(* IEC 61131-3 sources: Elmo_Master/Lasal_PRG/Welcon8Axis_EtherCAT_Test_With_RobotAxis/Network/TCPComNet, 1 file *)

(* ---- ONE_TCPComNet_Table.st ---- *)
#define OBJECTS_CONFIG

#include "..\..\Class\DataManager\DataManager.h"
//Define part of class DataManagerFIFO
#define MEMORY_Mark_DataMngFiFo    8
#include <.\lsl_st_mt.h>
#include "..\..\Class\TCPCommunication\TCPCommunication.h"
#include "..\..\Class\TCPCommunication\SalamanderDelay.h"

FUNCTION GLOBAL TAB ONE_TCPComNet
-1$UINT, 0$UINT,
0$UINT, 0$UINT,

15$UDINT,
TO_UDINT(916194998), "_CheckSum", 1$UINT, 0$UINT, 1$UINT,
TO_UDINT(3238142347), "_SigTCPComReceive", 1$UINT, 1$UINT, 0$UINT,
TO_UDINT(969826267), "_SigTCPDataManager", 1$UINT, 1$UINT, 1$UINT,
TO_UDINT(794617671), "CriticalSection", 0$UINT, 4$UINT, 10$UINT,
TO_UDINT(4008337867), "DataManager", 1$UINT, 1$UINT, 0$UINT,
TO_UDINT(2873804345), "DataManagerFIFO", 1$UINT, 1$UINT, 10$UINT,
TO_UDINT(2393054465), "DataManagerPriority", 1$UINT, 0$UINT, 1$UINT,
TO_UDINT(2602835227), "GetTaskHandle", 0$UINT, 2$UINT, 1$UINT,
TO_UDINT(2225119864), "MerkerEx", 1$UINT, 22$UINT, 2$UINT,
TO_UDINT(3534980377), "RamRingBuffer", 1$UINT, 1$UINT, 1$UINT,
TO_UDINT(1850111279), "String", 1$UINT, 11$UINT, 1$UINT,
TO_UDINT(2898603620), "StringInternal", 1$UINT, 86$UINT, 0$UINT,
TO_UDINT(4051501096), "TCP_MotionIF_Dummy", 0$UINT, 0$UINT, 1$UINT,
TO_UDINT(3704218787), "TCPCommunication", 1$UINT, 20$UINT, 1$UINT,
TO_UDINT(3232495061), "VirtualBaseInit", 1$UINT, 3$UINT, 0$UINT,

1$UINT, TO_UDINT(4103985232), "_SIGTCPDATAMANAGER1\TCPCOMMUNICATION\CHECKSUM",

_NO_ATTR, TO_UDINT(2464426676), "_SIGTCPDATAMANAGER1",

1$UINT, TO_UDINT(3019548784), "_SIGTCPDATAMANAGER1\_BASE\DATAMANAGERPRIORITY\DATAMANAGERFIFO_PRIO0\SECTION",
1$UINT, TO_UDINT(2759965747), "_SIGTCPDATAMANAGER1\_BASE\DATAMANAGERPRIORITY\DATAMANAGERFIFO_PRIO1\SECTION",
1$UINT, TO_UDINT(2634842358), "_SIGTCPDATAMANAGER1\_BASE\DATAMANAGERPRIORITY\DATAMANAGERFIFO_PRIO2\SECTION",
1$UINT, TO_UDINT(2323092661), "_SIGTCPDATAMANAGER1\_BASE\DATAMANAGERPRIORITY\DATAMANAGERFIFO_PRIO3\SECTION",
1$UINT, TO_UDINT(3994483068), "_SIGTCPDATAMANAGER1\_BASE\DATAMANAGERPRIORITY\DATAMANAGERFIFO_PRIO4\SECTION",
1$UINT, TO_UDINT(4184730943), "_SIGTCPDATAMANAGER1\_BASE\DATAMANAGERPRIORITY\DATAMANAGERFIFO_PRIO5\SECTION",
1$UINT, TO_UDINT(3235959290), "_SIGTCPDATAMANAGER1\_BASE\DATAMANAGERPRIORITY\DATAMANAGERFIFO_PRIO6\SECTION",
1$UINT, TO_UDINT(3617310137), "_SIGTCPDATAMANAGER1\_BASE\DATAMANAGERPRIORITY\DATAMANAGERFIFO_PRIO7\SECTION",
1$UINT, TO_UDINT(136448616), "_SIGTCPDATAMANAGER1\_BASE\DATAMANAGERPRIORITY\DATAMANAGERFIFO_PRIO8\SECTION",
1$UINT, TO_UDINT(525934123), "_SIGTCPDATAMANAGER1\_BASE\DATAMANAGERPRIORITY\DATAMANAGERFIFO_PRIO9\SECTION",

1$UINT, TO_UDINT(1713339845), "_SIGTCPDATAMANAGER1\_BASE\DATAMANAGERPRIORITY\DATAMANAGERFIFO_PRIO0",
1$UINT, TO_UDINT(286805331), "_SIGTCPDATAMANAGER1\_BASE\DATAMANAGERPRIORITY\DATAMANAGERFIFO_PRIO1",
1$UINT, TO_UDINT(2282822889), "_SIGTCPDATAMANAGER1\_BASE\DATAMANAGERPRIORITY\DATAMANAGERFIFO_PRIO2",
1$UINT, TO_UDINT(4279643263), "_SIGTCPDATAMANAGER1\_BASE\DATAMANAGERPRIORITY\DATAMANAGERFIFO_PRIO3",
1$UINT, TO_UDINT(1634908636), "_SIGTCPDATAMANAGER1\_BASE\DATAMANAGERPRIORITY\DATAMANAGERFIFO_PRIO4",
1$UINT, TO_UDINT(376801610), "_SIGTCPDATAMANAGER1\_BASE\DATAMANAGERPRIORITY\DATAMANAGERFIFO_PRIO5",
1$UINT, TO_UDINT(2407323888), "_SIGTCPDATAMANAGER1\_BASE\DATAMANAGERPRIORITY\DATAMANAGERFIFO_PRIO6",
1$UINT, TO_UDINT(4168869990), "_SIGTCPDATAMANAGER1\_BASE\DATAMANAGERPRIORITY\DATAMANAGERFIFO_PRIO7",
1$UINT, TO_UDINT(1757738487), "_SIGTCPDATAMANAGER1\_BASE\DATAMANAGERPRIORITY\DATAMANAGERFIFO_PRIO8",
1$UINT, TO_UDINT(532923745), "_SIGTCPDATAMANAGER1\_BASE\DATAMANAGERPRIORITY\DATAMANAGERFIFO_PRIO9",

1$UINT, TO_UDINT(3843458400), "_SIGTCPDATAMANAGER1\_BASE\DATAMANAGERPRIORITY",

1$UINT, TO_UDINT(1596713124), "_SIGTCPDATAMANAGER1\_BASE\DATAMNGGETTASKHANDLE1",

1$UINT, TO_UDINT(2770825344), "_SIGTCPDATAMANAGER1\TCPCOMMUNICATION\RAMRINGMERKEREX",
1$UINT, TO_UDINT(450202565), "_SIGTCPDATAMANAGER1\TCPCOMMUNICATION\THREADNAME\MERKEREX0",

1$UINT, TO_UDINT(3841123865), "_SIGTCPDATAMANAGER1\TCPCOMMUNICATION\RAMRINGBUFFER",

1$UINT, TO_UDINT(495891216), "_SIGTCPDATAMANAGER1\TCPCOMMUNICATION\THREADNAME",

_NO_ATTR, TO_UDINT(3063429709), "TCP_MOTIONIF_DUMMY1",

1$UINT, TO_UDINT(3070397306), "_SIGTCPDATAMANAGER1\TCPCOMMUNICATION",

//Internal connections
0$UDINT,
28$UDINT,
TO_UDINT(1), "DataMngGetTaskHandle1", TO_UDINT(23),
TO_UDINT(1), "DataManagerPriority", TO_UDINT(22),
TO_UDINT(1), "TCPCommunication", TO_UDINT(29),
TO_UDINT(12), "Section", TO_UDINT(2),
TO_UDINT(13), "Section", TO_UDINT(3),
TO_UDINT(14), "Section", TO_UDINT(4),
TO_UDINT(15), "Section", TO_UDINT(5),
TO_UDINT(16), "Section", TO_UDINT(6),
TO_UDINT(17), "Section", TO_UDINT(7),
TO_UDINT(18), "Section", TO_UDINT(8),
TO_UDINT(19), "Section", TO_UDINT(9),
TO_UDINT(20), "Section", TO_UDINT(10),
TO_UDINT(21), "Section", TO_UDINT(11),
TO_UDINT(22), "DataManagerFiFo_Prio0", TO_UDINT(12),
TO_UDINT(22), "DataManagerFiFo_Prio1", TO_UDINT(13),
TO_UDINT(22), "DataManagerFiFo_Prio2", TO_UDINT(14),
TO_UDINT(22), "DataManagerFiFo_Prio3", TO_UDINT(15),
TO_UDINT(22), "DataManagerFiFo_Prio4", TO_UDINT(16),
TO_UDINT(22), "DataManagerFiFo_Prio5", TO_UDINT(17),
TO_UDINT(22), "DataManagerFiFo_Prio6", TO_UDINT(18),
TO_UDINT(22), "DataManagerFiFo_Prio7", TO_UDINT(19),
TO_UDINT(22), "DataManagerFiFo_Prio8", TO_UDINT(20),
TO_UDINT(22), "DataManagerFiFo_Prio9", TO_UDINT(21),
TO_UDINT(27), "MerkerEx0", TO_UDINT(25),
TO_UDINT(29), "RamRingBuffer", TO_UDINT(26),
TO_UDINT(29), "RamRingMerkerEx", TO_UDINT(24),
TO_UDINT(29), "CheckSum", TO_UDINT(0),
TO_UDINT(29), "ThreadName", TO_UDINT(27),
0$UDINT,
5$UDINT,
TO_UDINT(1), "coTCPCommunication", TO_UDINT(29), "ClassSvr",
TO_UDINT(26), "Data", TO_UDINT(24), "m_udLength",
TO_UDINT(27), "DataBuffer", TO_UDINT(25), "m_udLength",
TO_UDINT(28), "_SigTCPDataManager", TO_UDINT(1), "ClassSvr",
TO_UDINT(29), "coDataMng", TO_UDINT(1), "ClassSvr",

//Initialization values
0$UDINT,
18$UDINT,
TO_UDINT(1), "AcceptOfflineJobs", TO_UDINT(1),//|TCPComNet._SigTCPDataManager1.AcceptOfflineJobs;
TO_UDINT(1), "ComPort", TO_UDINT(500),//|TCPComNet._SigTCPDataManager1.ComPort;
TO_UDINT(1), "LogEnable", TO_UDINT(0),//|TCPComNet._SigTCPDataManager1.LogEnable;
TO_UDINT(1), "DeactivateCom", TO_UDINT(0),//|TCPComNet._SigTCPDataManager1.DeactivateCom;
TO_UDINT(1), "LogFilter", TO_UDINT(0),//|TCPComNet._SigTCPDataManager1.LogFilter;
TO_UDINT(1), "SizeOfComBuffers", TO_UDINT(100 kB),//|TCPComNet._SigTCPDataManager1.SizeOfComBuffers;
TO_UDINT(1), "SizeOfComBufferRecv", TO_UDINT(100 kB),//|TCPComNet._SigTCPDataManager1.SizeOfComBufferRecv;
TO_UDINT(24), "ThreadSafe", TO_UDINT(0),//|TCPComNet.TCPCommunication\_SigTCPDataManager1\RamRingMerkerEx.ThreadSafe;
TO_UDINT(25), "ThreadSafe", TO_UDINT(0),//|TCPComNet.ThreadName\TCPCommunication\_SigTCPDataManager1\MerkerEx0.ThreadSafe;
TO_UDINT(27), "SingleRealloc", TO_UDINT(1),//|TCPComNet.TCPCommunication\_SigTCPDataManager1\ThreadName.SingleRealloc;
TO_UDINT(28), "SourceID", TO_UDINT(1),//|TCPComNet.TCP_MotionIF_Dummy1.SourceID;
TO_UDINT(28), "MotionControlIF", TO_UDINT(0),//|TCPComNet.TCP_MotionIF_Dummy1.MotionControlIF;
TO_UDINT(29), "ComPort", TO_UDINT(500),//|TCPComNet._SigTCPDataManager1\TCPCommunication.ComPort;
TO_UDINT(29), "LogEnable", TO_UDINT(0),//|TCPComNet._SigTCPDataManager1\TCPCommunication.LogEnable;
TO_UDINT(29), "DeactivateCom", TO_UDINT(0),//|TCPComNet._SigTCPDataManager1\TCPCommunication.DeactivateCom;
TO_UDINT(29), "coLogFilter", TO_UDINT(0),//|TCPComNet._SigTCPDataManager1\TCPCommunication.coLogFilter;
TO_UDINT(29), "SizeOfComBuffers", TO_UDINT(100 kB),//|TCPComNet._SigTCPDataManager1\TCPCommunication.SizeOfComBuffers;
TO_UDINT(29), "SizeOfComBufferRecv", TO_UDINT(100 kB),//|TCPComNet._SigTCPDataManager1\TCPCommunication.SizeOfComBufferRecv;

//Symbolic initialization values
0$UDINT,
0$UDINT,

//Initialization of string values
0$UDINT,
0$UDINT,

//Configuration of tasks (RealTime, Cyclic, Background)
0$UDINT,
1$UDINT,
TO_UDINT(23), (1000)$UDINT, 4194303$DINT, 	//_SIGTCPDATAMANAGER1\_BASE\DATAMNGGETTASKHANDLE1

0$UDINT,
2$UDINT,
TO_UDINT(1), (10)$UDINT, 4194303$DINT, 	//_SIGTCPDATAMANAGER1
TO_UDINT(23), (1000)$UDINT, 4194303$DINT, 	//_SIGTCPDATAMANAGER1\_BASE\DATAMNGGETTASKHANDLE1

0$UDINT,
1$UDINT,
TO_UDINT(23), (1000)$UDINT, 4194303$DINT, 	//_SIGTCPDATAMANAGER1\_BASE\DATAMNGGETTASKHANDLE1

//External connections
0$UDINT,
0$UDINT,

//Magic internal connections
0$UDINT,
7$UDINT,
TO_UDINT(29), "coIntern", TO_UDINT(1), "InternConnection",
TO_UDINT(29), "coIpToConnect", TO_UDINT(1), "IPtoConnect",
TO_UDINT(29), "coStationToConnect", TO_UDINT(1), "StationToConnect",
TO_UDINT(29), "coLogFilter", TO_UDINT(1), "LogFilter",
TO_UDINT(29), "ErrRuntime", TO_UDINT(1), "ErrRuntime",
TO_UDINT(29), "SizeOfComBuffers", TO_UDINT(1), "SizeOfComBuffers",
TO_UDINT(29), "SizeOfComBufferRecv", TO_UDINT(1), "SizeOfComBufferRecv",

//Configuration of timeslots of tasks (RealTime, Cyclic)
#ifdef __LSLLDR_TIMESLOTS__
0$UDINT,
0$UDINT,

0$UDINT,
0$UDINT,

#endif //__LSLLDR_TIMESLOTS__

//MultiMaster connections
#ifdef __LSLLDR_MULTIMASTER__
0$UDINT,
0$UDINT,
#endif //__LSLLDR_MULTIMASTER__

//Configuration for task ID (RealTime, CyclicTime)
#ifdef __LSLLDR_TASKID__
"\\\\TASKS2  "
0$UDINT,
1$UDINT,
(0)$UDINT, 	//_SIGTCPDATAMANAGER1\_BASE\DATAMNGGETTASKHANDLE1

0$UDINT,
2$UDINT,
(0)$UDINT, 	//_SIGTCPDATAMANAGER1
(0)$UDINT, 	//_SIGTCPDATAMANAGER1\_BASE\DATAMNGGETTASKHANDLE1

0$UDINT,
1$UDINT,
(0)$UDINT, 	//_SIGTCPDATAMANAGER1\_BASE\DATAMNGGETTASKHANDLE1

#endif //__LSLLDR_TASKID__

END_FUNCTION
